// TIA Portal project "OTOMATIK ETIKETLEME MAKINESI UYGULAMASI" (V18)

(* hardware
DEVICE "S7-1200 station_1"  S7-1200 Station
   slot 0: "Rack_0"  S7-1200 Rack  Rack  V1.0
   slot 1: "PLC_1"  CPU 1214C AC/DC/Rly  6ES7 214-1BG40-0XB0  V4.6
*)

// ===== PLC "PLC_1"  CPU 1214C AC/DC/Rly =====

VAR_GLOBAL   // PLC tag table "Default tag table"
   "START BUT" AT %I0.0 : Bool;
   "STOP BUT" AT %I0.1 : Bool;
   "YUKARIDA SENSORU" AT %I0.2 : Bool;
   "ASAGIDA SENSORU" AT %I0.3 : Bool;
   "VALF ASAGI" AT %Q0.0 : Bool;
   "VALF YUKARI" AT %Q0.1 : Bool;
   "SISTEM START MEM" AT %M10.0 : Bool;
END_VAR

// folder: System blocks/Program resources

DATA_BLOCK "TIMER 1"   // DB1
{ S7_Optimized_Access := 'TRUE' }
AUTHOR : Simatic
FAMILY : IEC
NAME : IEC_TMR
VERSION : 1.0
// stored: InstanceOfName IEC_TIMER
"IEC_TIMER"
BEGIN
END_DATA_BLOCK

// folder: (top level)

ORGANIZATION_BLOCK "Main"   // OB1, LAD, ProgramCycle
TITLE = "Main Program Sweep (Cycle)"
{ S7_Optimized_Access := 'TRUE' }
VERSION : 0.1
   VAR_INPUT
      Initial_Call : Bool;   // Initial call of this OB
      Remanence : Bool;   // =True, if remanent data are available
   END_VAR
BEGIN

REGION Network 1: SISTEM GENEL START
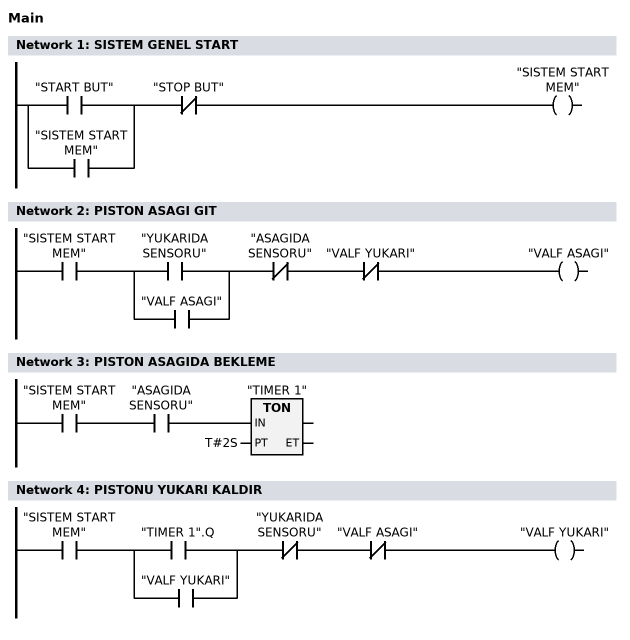
   RUNG wire#powerrail
      Contact( "START BUT" )
      wire#w1
      I_Contact( "STOP BUT" )
      Coil( "SISTEM START MEM" )
   END_RUNG
   RUNG wire#powerrail
      Contact( "SISTEM START MEM" )
   END_RUNG wire#w1
   // the same network as SCL:
   "SISTEM START MEM" := ("START BUT" OR "SISTEM START MEM") AND NOT "STOP BUT";
END_REGION

REGION Network 2: PISTON ASAGI GIT
   RUNG wire#powerrail
      Contact( "SISTEM START MEM" )
      wire#w1
      Contact( "YUKARIDA SENSORU" )
      wire#w2
      I_Contact( "ASAGIDA SENSORU" )
      I_Contact( "VALF YUKARI" )
      Coil( "VALF ASAGI" )
   END_RUNG
   RUNG wire#w1
      Contact( "VALF ASAGI" )
   END_RUNG wire#w2
   // the same network as SCL:
   "VALF ASAGI" := "SISTEM START MEM" AND ("YUKARIDA SENSORU" OR "VALF ASAGI") AND NOT "ASAGIDA SENSORU" AND NOT "VALF YUKARI";
END_REGION

REGION Network 3: PISTON ASAGIDA BEKLEME
   "TIMER 1".TON(IN := "SISTEM START MEM" AND "ASAGIDA SENSORU", PT := T#2S);
END_REGION

REGION Network 4: PISTONU YUKARI KALDIR
   RUNG wire#powerrail
      Contact( "SISTEM START MEM" )
      wire#w1
      Contact( "TIMER 1".Q )
      wire#w2
      I_Contact( "YUKARIDA SENSORU" )
      I_Contact( "VALF ASAGI" )
      Coil( "VALF YUKARI" )
   END_RUNG
   RUNG wire#w1
      Contact( "VALF YUKARI" )
   END_RUNG wire#w2
   // the same network as SCL:
   "VALF YUKARI" := "SISTEM START MEM" AND ("TIMER 1".Q OR "VALF YUKARI") AND NOT "YUKARIDA SENSORU" AND NOT "VALF ASAGI";
END_REGION
END_ORGANIZATION_BLOCK